Fanuc KAREL source: KT00745.KL

PROGRAM KT00745
%NOLOCKGROUP
VAR
  ARG: ARRAY[4] OF XYZWPR
  OUT: INTEGER
BEGIN
  OUT = ARRAY_LEN(ARG)
END KT00745
